Fanuc KAREL source: KA00171.KL

PROGRAM KA00171
%NOLOCKGROUP
VAR
  SRC: ARRAY[4] OF BOOLEAN
  DST: ARRAY[4] OF JOINTPOS
BEGIN
  DST = SRC
END KA00171
